// TwinCAT 3 PLC project ExamplePLC
// ProgramVersion: 3.1.4024.0
// libraries:
//   MachineLibrary, * (PLC-Template)
//   Tc2_Standard, * (Beckhoff Automation GmbH)
//   Tc2_System, * (Beckhoff Automation GmbH)
//   Tc2_Utilities, * (Beckhoff Automation GmbH)
//   Tc3_IotBase, * (Beckhoff Automation GmbH)
//   Tc3_JsonXml, * (Beckhoff Automation GmbH)
//   Tc3_Module, * (Beckhoff Automation GmbH)
//   MachineLibrary, * (PLC-Template)
// project tree:
//   Communication/MQTT/_DUTs/ ST_MqttConfiguration.TcDUT, ST_MqttStatus.TcDUT
//   Communication/MQTT/ FB_MqttStatePublisher.TcPOU
//   / PlcTask.TcTTO
//   POUs/ FB_Machine.TcPOU, MAIN.TcPOU
//   Stations/ExampleStation/_DUTs/ ST_ExampleStationConfiguration.TcDUT, ST_ExampleStationStatus.TcDUT
//   Stations/ExampleStation/_ENUMs/ E_ExampleStationRunStep.TcDUT
//   Stations/ExampleStation/ FB_ExampleStation.TcPOU
//   Simulation/SoftwareSim/_DUTs/ ST_ExampleSoftwareSimConfiguration.TcDUT, ST_ExampleSoftwareSimStatus.TcDUT
//   Simulation/SoftwareSim/_ENUMs/ E_ExampleSoftwareSimStep.TcDUT
//   Simulation/SoftwareSim/ FB_ExampleSoftwareSim.TcPOU
//   Stations/ExampleStation/Transaction/_DUTs/ ST_ExampleRequest.TcDUT, ST_ExampleResponse.TcDUT
//   Stations/ExampleStation/Transaction/ FB_ExampleTransaction.TcPOU
//   Simulation/DosingProcessSim/_DUTs/ ST_DosingProcessSimConfiguration.TcDUT, ST_DosingProcessSimStatus.TcDUT
//   Simulation/DosingProcessSim/ FB_DosingProcessSim.TcPOU
//   Stations/DosingStation/_DUTs/ ST_DosingStationConfiguration.TcDUT, ST_DosingStationStatus.TcDUT
//   Stations/DosingStation/ FB_DosingStation.TcPOU
// real-time tasks:
//   TASK PlcTask: cycle T#10ms, priority 20, ADS port 350

CONFIGURATION ExamplePLC
    RESOURCE PLC ON TwinCAT3
        TASK PlcTask(INTERVAL := T#10ms, PRIORITY := 20);
        PROGRAM MAIN WITH PlcTask : MAIN;
    END_RESOURCE
END_CONFIGURATION

// ---- Communication/MQTT/_DUTs/ST_MqttConfiguration.TcDUT
TYPE ST_MqttConfiguration :
STRUCT
	enable					: BOOL := TRUE; //connect to the broker and publish state
	hostName				: STRING(255) := 'broker.hivemq.com'; //public test broker, replace with your own
	hostPort				: UINT := 1883; //8883 for TLS
	stateTopic				: STRING(255) := 'plc-template/example/state'; //machine state is published here as JSON
	commandTopic			: STRING(255) := 'plc-template/example/cmd'; //START, STOP or RESET
	enableRemoteCommands	: BOOL := FALSE; //accept commands on commandTopic. Off by default: anyone on a public broker can publish to it
	publishInterval			: TIME := T#10S; //state is also published on every state change
END_STRUCT
END_TYPE

// ---- Communication/MQTT/_DUTs/ST_MqttStatus.TcDUT
TYPE ST_MqttStatus :
STRUCT
	connected				: BOOL; //connected to the broker
	subscribed				: BOOL; //subscribed to commandTopic
	error					: BOOL; //client error
	errorCode				: HRESULT; //client error code
	publishCount			: UDINT; //messages published
	lastPayloadIn			: STRING(255); //last payload received on commandTopic
END_STRUCT
END_TYPE

// ---- Stations/ExampleStation/_DUTs/ST_ExampleStationConfiguration.TcDUT
TYPE ST_ExampleStationConfiguration :
STRUCT
	cycleDwell			: TIME := T#2S; //wait time between jobs while running
	maxCloseDwell		: TIME := T#10S; //longest closeDwell accepted in a request
END_STRUCT
END_TYPE

// ---- Stations/ExampleStation/_DUTs/ST_ExampleStationStatus.TcDUT
TYPE ST_ExampleStationStatus :
STRUCT
	runStep				: E_ExampleStationRunStep := E_ExampleStationRunStep.Idle; //running sequence step
	allOpen				: BOOL; //both actuators at home (open)
	allClosed			: BOOL; //both actuators at work (closed)
	
	job					: ST_ExampleRequest; //job being worked on
	cycleCount			: UDINT; //completed jobs
	lastCycleTime		: TIME; //duration of the last close/hold/open cycle
	jobsRejected		: UDINT; //requests rejected as invalid
	lastRejectText		: T_MaxString; //reason for the last rejection
	commError			: BOOL; //transaction timed out waiting for the software
END_STRUCT
END_TYPE

// ---- Stations/ExampleStation/_ENUMs/E_ExampleStationRunStep.TcDUT
{attribute 'qualified_only'}
{attribute 'strict'}
{attribute 'to_string'}
TYPE E_ExampleStationRunStep :
(
	Idle			:= 0, //not running
	RequestJob		:= 10, //raise attention, ask the software for a job
	WaitJob			:= 20, //wait for the request, validate it, ack or reject
	WaitWorking		:= 30, //wait for the software to drop trigger
	Close			:= 40, //closing both actuators
	HoldClosed		:= 50, //holding closed for the requested closeDwell
	Open			:= 60, //opening both actuators
	Report			:= 70, //send the response with tell
	WaitReportAck	:= 80, //wait for the software to acknowledge the response
	Dwell			:= 90 //wait before requesting the next job
);
END_TYPE

// ---- Simulation/SoftwareSim/_DUTs/ST_ExampleSoftwareSimConfiguration.TcDUT
TYPE ST_ExampleSoftwareSimConfiguration :
STRUCT
	enable				: BOOL := TRUE; //answer the station's transactions
	responseDelay		: TIME := T#500MS; //delay before each software action
	closeDwell			: TIME := T#1S; //closeDwell sent in each request
	
	//Fault injection
	freeze				: BOOL; //stop responding where it is (tests the commTimeout)
	sendInvalidRequest	: BOOL; //send closeDwell = T#0S (station should reject it)
END_STRUCT
END_TYPE

// ---- Simulation/SoftwareSim/_DUTs/ST_ExampleSoftwareSimStatus.TcDUT
TYPE ST_ExampleSoftwareSimStatus :
STRUCT
	step				: E_ExampleSoftwareSimStep := E_ExampleSoftwareSimStep.Idle; //current step
	requestsSent		: UDINT; //requests sent (trigger raised)
	responsesReceived	: UDINT; //responses received (tell acknowledged)
	aborts				: UDINT; //transactions aborted by the PLC
	lastResponse		: ST_ExampleResponse; //last response read on tell
END_STRUCT
END_TYPE

// ---- Simulation/SoftwareSim/_ENUMs/E_ExampleSoftwareSimStep.TcDUT
{attribute 'qualified_only'}
{attribute 'strict'}
{attribute 'to_string'}
TYPE E_ExampleSoftwareSimStep :
(
	Idle			:= 0, //waiting for attention
	SendTrigger		:= 10, //delay, then raise trigger with a request
	WaitTriggerAck	:= 20, //waiting for trigger_ack
	DropTrigger		:= 30, //delay, then drop trigger
	WaitTell		:= 40, //waiting for tell
	SendTellAck		:= 50, //delay, read response, raise tell_ack
	WaitTellDrop	:= 60, //waiting for tell to drop
	DropTellAck		:= 70 //drop tell_ack, transaction closed
);
END_TYPE

// ---- Stations/ExampleStation/Transaction/_DUTs/ST_ExampleRequest.TcDUT
(* Request from the software to the station, sent with trigger. *)
TYPE ST_ExampleRequest :
STRUCT
	cycleId				: UDINT; //id chosen by the software, echoed back in the response
	closeDwell			: TIME; //how long to hold the actuators closed
END_STRUCT
END_TYPE

// ---- Stations/ExampleStation/Transaction/_DUTs/ST_ExampleResponse.TcDUT
(* Response from the station to the software, sent with tell. *)
TYPE ST_ExampleResponse :
STRUCT
	cycleId				: UDINT; //cycleId from the request
	cycleTime			: TIME; //time to close, hold and open
	ok					: BOOL; //cycle completed without faults
END_STRUCT
END_TYPE

// ---- Simulation/DosingProcessSim/_DUTs/ST_DosingProcessSimConfiguration.TcDUT
TYPE ST_DosingProcessSimConfiguration :
STRUCT
	enable				: BOOL := TRUE; //simulate the flows (turn off when real I/O is linked)
	mainFlowBase		: LREAL := 200; //average main flow in l/min (set below 50 to test the low-low interlock)
	mainFlowSwing		: LREAL := 50; //main flow varies +/- this much in l/min
	swingPeriod			: TIME := T#60S; //period of the main flow variation, T#0S = constant
	maxDosingFlow		: LREAL := 80; //dosing flow at 100 % valve in l/min
	processLag			: TIME := T#2S; //time constant from valve position to dosing flow
END_STRUCT
END_TYPE

// ---- Simulation/DosingProcessSim/_DUTs/ST_DosingProcessSimStatus.TcDUT
TYPE ST_DosingProcessSimStatus :
STRUCT
	mainFlow			: LREAL; //simulated main flow in l/min
	dosingFlow			: LREAL; //simulated dosing flow in l/min
END_STRUCT
END_TYPE

// ---- Stations/DosingStation/_DUTs/ST_DosingStationConfiguration.TcDUT
TYPE ST_DosingStationConfiguration :
STRUCT
	ratio				: LREAL := 0.2; //dosing flow / main flow while running
END_STRUCT
END_TYPE

// ---- Stations/DosingStation/_DUTs/ST_DosingStationStatus.TcDUT
TYPE ST_DosingStationStatus :
STRUCT
	dosing				: BOOL; //PID in ratio control
	mainFlow			: LREAL; //main flow in l/min
	dosingFlow			: LREAL; //dosing flow in l/min
	dosingSetpoint		: LREAL; //dosing flow setpoint from the ratio, in l/min
	ratioActual			: LREAL; //dosing flow / main flow
	valvePosition		: LREAL; //dosing valve position in %
	mainFlowLow			: BOOL; //main flow below its low-low limit: dosing valve interlocked closed
END_STRUCT
END_TYPE

// ---- POUs/MAIN.TcPOU
PROGRAM MAIN
VAR
	{attribute 'OPC.UA.DA' := '1'}
	machine		: FB_Machine; //top-level module, start/stop with machine.ocmd
	
	(* Test harness
	----------------------------------------------------------------------------------------------------*)
	{attribute 'OPC.UA.DA' := '1'}
	softwareSim	: FB_ExampleSoftwareSim; //plays the software side of the station's trigger/tell
	{attribute 'OPC.UA.DA' := '1'}
	dosingSim	: FB_DosingProcessSim; //simulates the dosing station's flows
END_VAR

machine();

//Outside world: answers the example station's job requests
softwareSim(transaction := machine.exampleStation.transaction);

//Process simulation for the dosing station (turn off with dosingSim.cfg.enable when I/O is linked)
dosingSim(station := machine.dosingStation);

END_PROGRAM

// ---- POUs/FB_Machine.TcPOU
FUNCTION_BLOCK FB_Machine EXTENDS FB_Module
(*
	Top-level module. Starting/stopping the machine starts/stops both stations.
	Start/stop/reset from the HMI with ocmd, or over MQTT (see cfgMqtt.enableRemoteCommands).
*)
VAR_INPUT
	(* Stations
	----------------------------------------------------------------------------------------------------*)
	{attribute 'OPC.UA.DA' := '1'}
	exampleStation		: FB_ExampleStation;
	{attribute 'OPC.UA.DA' := '1'}
	dosingStation		: FB_DosingStation; //ratio control loop example
	
	(* Communication
	----------------------------------------------------------------------------------------------------*)
	{attribute 'OPC.UA.DA' := '1'}
	{attribute 'OPC.UA.DA.StructuredType' := '1'}
	cfgMqtt				: ST_MqttConfiguration; //MQTT configuration
END_VAR
VAR
	{attribute 'OPC.UA.DA' := '0'} // internal MQTT client holds pointers OPC UA can't publish; status is in cfgMqtt/dashboard
	mqtt				: FB_MqttStatePublisher; //MQTT state publisher
END_VAR

SUPER^();

Stations();
Permissives();
Communication();

METHOD PROTECTED Communication
mqtt(cfg 			:= cfgMqtt,
	 machineState 	:= sts.State,
	 cycleCount 	:= exampleStation.stsStation.cycleCount);

//Remote commands are handled like program commands
IF mqtt.cmd <> E_ModuleCommand.None THEN
	pcmd := mqtt.cmd;
END_IF
END_METHOD

METHOD PROTECTED Permissives //set module permissives and interlocks
//Started once every station is running
PermStartComplete.cfg.condText[0] := 'Example station started';
PermStartComplete.cfg.condText[1] := 'Dosing station started';
PermStartComplete.perm.0 := exampleStation.sts.Started;
PermStartComplete.perm.1 := dosingStation.sts.Started;

//Stopped once every station is stopped
PermStopComplete.cfg.condText[0] := 'Example station stopped';
PermStopComplete.cfg.condText[1] := 'Dosing station stopped';
PermStopComplete.perm.0 := exampleStation.sts.Stopped;
PermStopComplete.perm.1 := dosingStation.sts.Stopped;

//A faulted station stops the machine
IntlkAuto.cfg.condText[0] := 'Example station not faulted';
IntlkAuto.cfg.condText[1] := 'Dosing station not faulted';
IntlkAuto.perm.0 := NOT exampleStation.sts.Faulted;
IntlkAuto.perm.1 := NOT dosingStation.sts.Faulted;
END_METHOD

METHOD PUBLIC Reset : BOOL
exampleStation.cmdReset := TRUE;
dosingStation.cmdReset := TRUE;
Reset := TRUE;
END_METHOD

METHOD PROTECTED Started : BOOL
//Stations run their own sequences while the machine is started
END_METHOD

METHOD PROTECTED Starting : BOOL
exampleStation.pcmd := E_ModuleCommand.Start;
dosingStation.pcmd := E_ModuleCommand.Start;
END_METHOD

METHOD PROTECTED Stations //call child modules
exampleStation();
dosingStation();

inpChildFaulted := exampleStation.sts.Faulted OR dosingStation.sts.Faulted;
END_METHOD

METHOD PROTECTED Stopping : BOOL
exampleStation.pcmd := E_ModuleCommand.Stop;
dosingStation.pcmd := E_ModuleCommand.Stop;
END_METHOD

END_FUNCTION_BLOCK

// ---- Stations/ExampleStation/FB_ExampleStation.TcPOU
FUNCTION_BLOCK FB_ExampleStation EXTENDS FB_Module
(*
	Example station with two 2-state actuators and a trigger/tell transaction.
	Home position = OPEN, Work position = CLOSED.
	
	Starting (homing)	: open both actuators, Started once both are open
	Started (running)	: one job per cycle:
						  ask the software for a job (attention), validate and ack the request,
						  close both, hold for request.closeDwell, open both, report (tell), dwell
	Stopping			: abort any open transaction, open both actuators (safe position)
	Stopped				: actuators follow operator commands (manual mode)
	
	The actuators are configured with no feedback so the example runs without hardware.
	Clear homeNoFdbk/workNoFdbk and link homeFdbk/workFdbk/outHome/outWork to use real I/O.
*)
VAR_INPUT
	{attribute 'OPC.UA.DA' := '1'}
	{attribute 'OPC.UA.DA.StructuredType' := '1'}
	cfg					: ST_ExampleStationConfiguration; //configuration
	
	(* Devices
	----------------------------------------------------------------------------------------------------*)
	{attribute 'OPC.UA.DA' := '1'}
	actuatorA			: FB_Actuator2State := (cfg := (actuatorId := 'Actuator A', homeNoFdbk := TRUE, workNoFdbk := TRUE));
	{attribute 'OPC.UA.DA' := '1'}
	actuatorB			: FB_Actuator2State := (cfg := (actuatorId := 'Actuator B', homeNoFdbk := TRUE, workNoFdbk := TRUE));
	
	(* Communication
	----------------------------------------------------------------------------------------------------*)
	{attribute 'OPC.UA.DA' := '1'}
	transaction			: FB_ExampleTransaction := (cfg := (commTimeout := T#10S)); //job request/response with the software
END_VAR
VAR_OUTPUT
	{attribute 'OPC.UA.DA' := '1'}
	{attribute 'OPC.UA.DA.Access' := '1'}
	{attribute 'OPC.UA.DA.StructuredType' := '1'}
	stsStation			: ST_ExampleStationStatus; //station specific status (module status is in sts)
END_VAR
VAR
	//Timers
	dwellTimer			: TON; //dwell between cycles
	holdTimer			: TON; //holds the actuators closed for job.closeDwell
	cycleTimer			: TON := (PT := T#1D); //measures one close/hold/open cycle
END_VAR

SUPER^();

Devices();
Permissives();
StatusOut();

METHOD PROTECTED CloseAll //command all actuators to work (closed)
IF NOT actuatorA.sts.atWork AND NOT actuatorA.sts.goingToWork THEN
	actuatorA.ToWork();
END_IF
IF NOT actuatorB.sts.atWork AND NOT actuatorB.sts.goingToWork THEN
	actuatorB.ToWork();
END_IF
END_METHOD

METHOD PROTECTED Devices //call child devices
//Devices follow this module's mode through childCtrl
actuatorA(parentCtrl := childCtrl);
actuatorB(parentCtrl := childCtrl);
transaction();

//Report child faults to the module
inpChildFaulted := actuatorA.fault.active OR actuatorB.fault.active;
END_METHOD

METHOD PROTECTED OpenAll //command all actuators to home (open)
IF NOT actuatorA.sts.atHome AND NOT actuatorA.sts.goingToHome THEN
	actuatorA.ToHome();
END_IF
IF NOT actuatorB.sts.atHome AND NOT actuatorB.sts.goingToHome THEN
	actuatorB.ToHome();
END_IF
END_METHOD

METHOD PROTECTED Permissives //set module permissives and interlocks
//Homing is complete when all actuators are open
PermStartComplete.cfg.condText[0] := 'Actuator A open';
PermStartComplete.cfg.condText[1] := 'Actuator B open';
PermStartComplete.perm.0 := actuatorA.sts.atHome;
PermStartComplete.perm.1 := actuatorB.sts.atHome;

//Stopping is complete when all actuators are open, or faulted so they cannot move
PermStopComplete.cfg.condText[0] := 'Actuator A open or faulted';
PermStopComplete.cfg.condText[1] := 'Actuator B open or faulted';
PermStopComplete.perm.0 := actuatorA.sts.atHome OR actuatorA.fault.active;
PermStopComplete.perm.1 := actuatorB.sts.atHome OR actuatorB.fault.active;

//A faulted actuator stops the station
IntlkAuto.cfg.condText[0] := 'Actuator A not faulted';
IntlkAuto.cfg.condText[1] := 'Actuator B not faulted';
IntlkAuto.perm.0 := NOT actuatorA.fault.active;
IntlkAuto.perm.1 := NOT actuatorB.fault.active;
END_METHOD

METHOD PUBLIC Reset : BOOL
actuatorA.Reset();
actuatorB.Reset();
transaction.Reset();
Reset := TRUE;
END_METHOD

METHOD PROTECTED Started : BOOL
//Running sequence: one trigger/tell transaction per close/open cycle
CASE stsStation.runStep OF
	
	E_ExampleStationRunStep.Idle:
		stsStation.runStep := E_ExampleStationRunStep.RequestJob;
		
	E_ExampleStationRunStep.RequestJob:
		IF transaction.sts.Idle THEN
			transaction.Start(); //raises attention
			stsStation.runStep := E_ExampleStationRunStep.WaitJob;
		END_IF
		
	E_ExampleStationRunStep.WaitJob:
		IF transaction.sts.Request_Start THEN
			IF ValidateJob(transaction.request) THEN
				stsStation.job := transaction.request;
				transaction.SetRequestACK();
				stsStation.runStep := E_ExampleStationRunStep.WaitWorking;
			ELSE
				transaction.Abort();
				stsStation.jobsRejected := stsStation.jobsRejected + 1;
				stsStation.runStep := E_ExampleStationRunStep.Dwell;
			END_IF
		END_IF
		
	E_ExampleStationRunStep.WaitWorking:
		IF transaction.sts.Working THEN
			stsStation.runStep := E_ExampleStationRunStep.Close;
		END_IF
		
	E_ExampleStationRunStep.Close:
		CloseAll();
		IF stsStation.allClosed THEN
			stsStation.runStep := E_ExampleStationRunStep.HoldClosed;
		END_IF
		
	E_ExampleStationRunStep.HoldClosed:
		IF holdTimer.Q THEN
			stsStation.runStep := E_ExampleStationRunStep.Open;
		END_IF
		
	E_ExampleStationRunStep.Open:
		OpenAll();
		IF stsStation.allOpen THEN
			stsStation.lastCycleTime := cycleTimer.ET;
			stsStation.runStep := E_ExampleStationRunStep.Report;
		END_IF
		
	E_ExampleStationRunStep.Report:
		transaction.response.cycleId 	:= stsStation.job.cycleId;
		transaction.response.cycleTime 	:= stsStation.lastCycleTime;
		transaction.response.ok 		:= NOT (actuatorA.fault.active OR actuatorB.fault.active);
		transaction.FinishWork(); //raises tell
		stsStation.cycleCount := stsStation.cycleCount + 1;
		stsStation.runStep := E_ExampleStationRunStep.WaitReportAck;
		
	E_ExampleStationRunStep.WaitReportAck:
		IF transaction.sts.Idle THEN
			stsStation.runStep := E_ExampleStationRunStep.Dwell;
		END_IF
		
	E_ExampleStationRunStep.Dwell:
		IF dwellTimer.Q THEN
			stsStation.runStep := E_ExampleStationRunStep.RequestJob;
		END_IF
		
END_CASE
END_METHOD

METHOD PROTECTED Starting : BOOL
//Homing: open all actuators, no transaction open
OpenAll();
AbortTransaction();
stsStation.runStep := E_ExampleStationRunStep.Idle;
END_METHOD

METHOD PROTECTED StatusOut //Set output status information
stsStation.allOpen 	:= actuatorA.sts.atHome AND actuatorB.sts.atHome;
stsStation.allClosed 	:= actuatorA.sts.atWork AND actuatorB.sts.atWork;

stsStation.commError 	:= transaction.sts.errTimeout;

//Monitoring timers
dwellTimer(IN := stsStation.runStep = E_ExampleStationRunStep.Dwell, PT := cfg.cycleDwell);
holdTimer(IN := stsStation.runStep = E_ExampleStationRunStep.HoldClosed, PT := stsStation.job.closeDwell);
cycleTimer(IN := stsStation.runStep = E_ExampleStationRunStep.Close
			OR stsStation.runStep = E_ExampleStationRunStep.HoldClosed
			OR stsStation.runStep = E_ExampleStationRunStep.Open);
END_METHOD

METHOD PROTECTED Stopping : BOOL
//Finish in the safe position: all actuators open, transaction closed
OpenAll();
AbortTransaction();
stsStation.runStep := E_ExampleStationRunStep.Idle;
END_METHOD

METHOD PROTECTED AbortTransaction //cancel an open transaction
IF transaction.sts.bBusy THEN
	transaction.Abort();
END_IF
END_METHOD

METHOD PROTECTED ValidateJob : BOOL //TRUE if the request can be worked on, sets lastRejectText otherwise
VAR_INPUT
	job			: ST_ExampleRequest;
END_VAR
IF job.closeDwell <= T#0S THEN
	stsStation.lastRejectText := 'closeDwell must be greater than 0';
ELSIF job.closeDwell > cfg.maxCloseDwell THEN
	stsStation.lastRejectText := 'closeDwell is longer than cfg.maxCloseDwell';
ELSE
	ValidateJob := TRUE;
	RETURN;
END_IF
ValidateJob := FALSE;
END_METHOD

END_FUNCTION_BLOCK

// ---- Stations/ExampleStation/Transaction/FB_ExampleTransaction.TcPOU
FUNCTION_BLOCK FB_ExampleTransaction EXTENDS FB_TriggerTell
(*
	Trigger/tell transaction for the example station, carrying ST_ExampleRequest in
	and ST_ExampleResponse out.
	
	FB_TriggerTell keeps its handshake bits internal. This FB is the transport layer:
	the software side writes trigger/tell_ack with WriteTrigger()/WriteTellAck() and
	reads the PLC bits from handshake. A real project would map these to OPC UA or MQTT.
*)
VAR_INPUT
	{attribute 'OPC.UA.DA' := '1'}
	{attribute 'OPC.UA.DA.StructuredType' := '1'}
	response			: ST_ExampleResponse; //set by the station before FinishWork()
END_VAR
VAR_OUTPUT
	{attribute 'OPC.UA.DA' := '1'}
	{attribute 'OPC.UA.DA.Access' := '1'}
	{attribute 'OPC.UA.DA.StructuredType' := '1'}
	request				: ST_ExampleRequest; //request latched when trigger rises
	{attribute 'OPC.UA.DA' := '1'}
	{attribute 'OPC.UA.DA.Access' := '1'}
	{attribute 'OPC.UA.DA.StructuredType' := '1'}
	handshake			: ST_TriggerTellHandshake; //copy of all handshake bits for the software side
END_VAR
VAR
	requestIn			: ST_ExampleRequest; //request written by the software with trigger
	
	//Oneshot triggers
	rtTrigger			: R_TRIG;
END_VAR

//Latch the request when the software raises trigger
rtTrigger(CLK := stHandshake.trigger);
IF rtTrigger.Q THEN
	request := requestIn;
END_IF

SUPER^();

handshake := stHandshake;

METHOD PUBLIC Response_Cleanup : BOOL //clear the response once the software acknowledged it
VAR
	emptyResponse : ST_ExampleResponse;
END_VAR
SUPER^.Response_Cleanup();
response := emptyResponse;
Response_Cleanup := TRUE;
END_METHOD

METHOD PUBLIC WriteTellAck //software side: set or clear tell_ack
VAR_INPUT
	value		: BOOL;
END_VAR
stHandshake.tell_ack := value;
END_METHOD

METHOD PUBLIC WriteTrigger //software side: set or clear trigger, with the request data
VAR_INPUT
	value		: BOOL;
	req			: ST_ExampleRequest; //only used when value is TRUE
END_VAR
IF value THEN
	requestIn := req;
END_IF
stHandshake.trigger := value;
END_METHOD

END_FUNCTION_BLOCK

// ---- Stations/DosingStation/FB_DosingStation.TcPOU
FUNCTION_BLOCK FB_DosingStation EXTENDS FB_Module
(*
	Example of a ratio control loop built from MachineLibrary blocks:
	
		flowMain (FB_AnalogInput)	main flow, the "wild" flow nobody controls
		flowDosing (FB_AnalogInput)	dosing flow, the process value
		dosingPid (FB_PID)			Ratio mode: dosing setpoint = cfg.ratio x main flow
		dosingValve					FB_ActuatorModulating driven by the PID output
	
	Starting	: PID off, valve closed
	Started		: PID in Ratio mode at cfg.ratio
	Stopping	: PID off, valve closed
	Interlock	: main flow low-low closes the valve (dosing into no flow is unsafe)
	
	No hardware needed: the valve has no position feedback (simulated stroke) and
	MAIN.dosingSim writes both flows into the analog inputs' simulation values.
	For real I/O, link flowMain.inpRaw, flowDosing.inpRaw and dosingValve.outRaw,
	and turn off MAIN.dosingSim.
*)
VAR_INPUT
	{attribute 'OPC.UA.DA' := '1'}
	{attribute 'OPC.UA.DA.StructuredType' := '1'}
	cfg					: ST_DosingStationConfiguration; //configuration
	
	(* Devices
	----------------------------------------------------------------------------------------------------*)
	{attribute 'OPC.UA.DA' := '1'}
	flowMain			: FB_AnalogInput := (cfg := (inputId := 'Main flow', units := 'l/min', euMax := 400, filterTime := T#500MS, limits := (LowLow := 50, Low := 100, High := 350, HighHigh := 380), alarmEnable := (lowLow := TRUE, low := TRUE, high := TRUE, highHigh := TRUE)));
	{attribute 'OPC.UA.DA' := '1'}
	flowDosing			: FB_AnalogInput := (cfg := (inputId := 'Dosing flow', units := 'l/min', euMax := 100, filterTime := T#500MS));
	{attribute 'OPC.UA.DA' := '1'}
	dosingPid			: FB_PID := (cfg := (loopId := 'Dosing', kp := 1.5, ti := T#3S, setpointMax := 100, ratioMax := 1, deviationEnable := TRUE, deviationLimit := 10));
	{attribute 'OPC.UA.DA' := '1'}
	dosingValve			: FB_ActuatorModulating := (cfg := (actuatorId := 'Dosing valve', noFdbk := TRUE, strokeTime := T#10S, failTimePositioning := T#30S));
END_VAR
VAR_OUTPUT
	{attribute 'OPC.UA.DA' := '1'}
	{attribute 'OPC.UA.DA.Access' := '1'}
	{attribute 'OPC.UA.DA.StructuredType' := '1'}
	stsStation			: ST_DosingStationStatus; //station specific status (module status is in sts)
END_VAR
VAR
END_VAR

SUPER^();

Devices();
Permissives();
StatusOut();

METHOD PROTECTED Devices //call child devices and connect the loop
//Inputs first, so the PID sees this scan's values
flowMain();
flowDosing();

dosingPid(pv		:= flowDosing.sts.value,
		  wildValue	:= flowMain.sts.value,
		  inpPvBad	:= NOT flowDosing.sts.valid,
		  parentCtrl := childCtrl);

//Dosing into a low main flow is not allowed: losing this closes the valve
dosingValve.intlk.cfg.condText[0] := 'Main flow not low-low';
dosingValve.intlk.perm.0 := NOT flowMain.sts.lowLow;
dosingValve(parentCtrl := childCtrl);

//PID output to the valve (program commands are only accepted in Auto)
IF dosingPid.sts.closedLoop AND dosingValve.sts.modeAuto THEN
	dosingValve.SetPosition(dosingPid.out);
END_IF

//Report child faults to the module
inpChildFaulted := dosingValve.fault.active OR dosingPid.fault.active
				OR flowMain.fault.active OR flowDosing.fault.active;
END_METHOD

METHOD PROTECTED Permissives //set module permissives and interlocks
//Homing is complete when the valve is closed and the loop is off
PermStartComplete.cfg.condText[0] := 'Dosing valve closed';
PermStartComplete.cfg.condText[1] := 'Dosing loop off';
PermStartComplete.perm.0 := dosingValve.sts.closed;
PermStartComplete.perm.1 := dosingPid.sts.loopMode = E_PIDLoopMode.Off;

//Stopping is complete when the valve is closed, or faulted so it cannot move
PermStopComplete.cfg.condText[0] := 'Dosing valve closed or faulted';
PermStopComplete.perm.0 := dosingValve.sts.closed OR dosingValve.fault.active;

//Faults stop the station
IntlkAuto.cfg.condText[0] := 'Dosing valve not faulted';
IntlkAuto.cfg.condText[1] := 'Dosing loop not faulted';
IntlkAuto.cfg.condText[2] := 'Flow signals good';
IntlkAuto.perm.0 := NOT dosingValve.fault.active;
IntlkAuto.perm.1 := NOT dosingPid.fault.active;
IntlkAuto.perm.2 := NOT (flowMain.fault.active OR flowDosing.fault.active);
END_METHOD

METHOD PUBLIC Reset : BOOL
flowMain.Reset();
flowDosing.Reset();
dosingPid.Reset();
dosingValve.Reset();
Reset := TRUE;
END_METHOD

METHOD PROTECTED Started : BOOL
//Running: ratio control. Re-issued when the ratio changes.
IF dosingPid.sts.loopMode <> E_PIDLoopMode.Ratio OR dosingPid.sts.ratio <> cfg.ratio THEN
	dosingPid.Ratio(cfg.ratio);
END_IF
END_METHOD

METHOD PROTECTED Starting : BOOL
//Homing: loop off, valve closed
SafeState();
END_METHOD

METHOD PROTECTED Stopping : BOOL
//Finish in the safe state: loop off, valve closed
SafeState();
END_METHOD

METHOD PROTECTED SafeState //loop off and valve closed
IF dosingPid.sts.loopMode <> E_PIDLoopMode.Off THEN
	dosingPid.Off();
END_IF
IF NOT dosingValve.sts.closed AND dosingValve.sts.setpoint <> dosingValve.cfg.minPosition THEN
	dosingValve.Close();
END_IF
END_METHOD

METHOD PROTECTED StatusOut //Set output status information
stsStation.dosing			:= dosingPid.sts.loopMode = E_PIDLoopMode.Ratio;
stsStation.mainFlow			:= flowMain.sts.value;
stsStation.dosingFlow		:= flowDosing.sts.value;
stsStation.dosingSetpoint	:= dosingPid.sts.setpoint;
stsStation.valvePosition	:= dosingValve.sts.position;
stsStation.mainFlowLow		:= flowMain.sts.lowLow;
IF flowMain.sts.value > 0 THEN
	stsStation.ratioActual := flowDosing.sts.value / flowMain.sts.value;
ELSE
	stsStation.ratioActual := 0;
END_IF
END_METHOD

END_FUNCTION_BLOCK

// ---- Communication/MQTT/FB_MqttStatePublisher.TcPOU
FUNCTION_BLOCK FB_MqttStatePublisher
(*
	Publishes the machine state as JSON over MQTT, and optionally accepts START/STOP/RESET.
	Shows how Tc3_IotBase and Tc3_JsonXml are used next to MachineLibrary.
	Payload example: {"state":"Started","cycleCount":12}
*)
VAR_INPUT
	{attribute 'OPC.UA.DA' := '1'}
	{attribute 'OPC.UA.DA.StructuredType' := '1'}
	cfg					: ST_MqttConfiguration; //configuration
	
	machineState		: E_ModuleState; //state to publish
	cycleCount			: UDINT; //cycle count to publish
END_VAR
VAR_OUTPUT
	cmd					: E_ModuleCommand; //remote command received this scan, None otherwise
	
	{attribute 'OPC.UA.DA' := '1'}
	{attribute 'OPC.UA.DA.Access' := '1'}
	{attribute 'OPC.UA.DA.StructuredType' := '1'}
	sts					: ST_MqttStatus;
END_VAR
VAR
	bInit				: BOOL := TRUE;
	
	//MQTT client
	client				: FB_IotMqttClient;
	queue				: FB_IotMqttMessageQueue;
	message				: FB_IotMqttMessage;
	
	//Publish
	json				: FB_JsonSaxWriter;
	stateText			: STRING;
	payloadOut			: STRING(255);
	publishRequest		: BOOL;
	machineStateLast	: E_ModuleState := E_ModuleState.Unknown;
	publishTimer		: TON;
	
	//Subscribe
	{attribute 'TcEncoding' := 'UTF-8'}
	topicIn				: STRING(255);
	{attribute 'TcEncoding' := 'UTF-8'}
	payloadIn			: STRING(255);
END_VAR

cmd := E_ModuleCommand.None;

IF NOT cfg.enable THEN
	sts.connected := sts.subscribed := FALSE;
	RETURN;
END_IF

IF bInit THEN
	Init();
	bInit := FALSE;
END_IF

Connection();
Publish();
Subscribe();

METHOD PROTECTED Connection //keep the client connected (must run every scan)
client.Execute(bConnect := TRUE);

sts.connected 	:= client.bConnected;
sts.error 		:= client.bError;
sts.errorCode 	:= client.hrErrorCode;
END_METHOD

METHOD PROTECTED Init : BOOL
client.sHostName 		:= cfg.hostName;
client.nHostPort 		:= cfg.hostPort;
client.ipMessageQueue 	:= queue; //route received messages into the queue
Init := TRUE;
END_METHOD

METHOD PROTECTED Publish //publish on state change and every publishInterval
publishTimer(IN := sts.connected AND NOT publishTimer.Q, PT := cfg.publishInterval);
publishRequest := publishRequest OR publishTimer.Q OR (machineState <> machineStateLast);
machineStateLast := machineState;

IF publishRequest AND sts.connected THEN
	stateText := TO_STRING(machineState);
	
	json.ResetDocument();
	json.StartObject();
	json.AddKey('state');
	json.AddString(stateText);
	json.AddKey('cycleCount');
	json.AddDint(UDINT_TO_DINT(cycleCount));
	json.EndObject();
	json.CopyDocument(payloadOut, SIZEOF(payloadOut));
	
	IF client.Publish(
		sTopic			:= cfg.stateTopic,
		pPayload		:= ADR(payloadOut),
		nPayloadSize	:= INT_TO_UDINT(LEN(payloadOut)),
		eQoS			:= TcIotMqttQos.AtMostOnceDelivery,
		bRetain			:= FALSE,
		bQueue			:= FALSE)
	THEN
		publishRequest := FALSE;
		sts.publishCount := sts.publishCount + 1;
	END_IF
END_IF
END_METHOD

METHOD PROTECTED Subscribe //receive remote commands
IF NOT cfg.enableRemoteCommands THEN
	RETURN;
END_IF

IF sts.connected AND NOT sts.subscribed THEN
	sts.subscribed := client.Subscribe(sTopic := cfg.commandTopic, eQoS := TcIotMqttQos.AtMostOnceDelivery);
ELSIF NOT sts.connected THEN
	sts.subscribed := FALSE;
END_IF

IF queue.nQueuedMessages > 0 THEN
	IF queue.Dequeue(fbMessage := message) THEN
		MEMSET(ADR(payloadIn), 0, SIZEOF(payloadIn));
		message.GetTopic(pTopic := ADR(topicIn), nTopicSize := SIZEOF(topicIn));
		message.GetPayload(pPayload := ADR(payloadIn), nPayloadSize := SIZEOF(payloadIn), bSetNullTermination := TRUE);
		sts.lastPayloadIn := payloadIn;
		
		IF payloadIn = 'START' THEN
			cmd := E_ModuleCommand.Start;
		ELSIF payloadIn = 'STOP' THEN
			cmd := E_ModuleCommand.Stop;
		ELSIF payloadIn = 'RESET' THEN
			cmd := E_ModuleCommand.Reset;
		END_IF
	END_IF
END_IF
END_METHOD

END_FUNCTION_BLOCK

// ---- Simulation/SoftwareSim/FB_ExampleSoftwareSim.TcPOU
FUNCTION_BLOCK FB_ExampleSoftwareSim
(*
	Plays the software (MES) side of FB_ExampleTransaction so the trigger/tell
	handshake can be tested without any outside software.
	
	For each transaction: wait for attention, send a request with trigger, drop trigger
	after trigger_ack, read the response on tell, acknowledge with tell_ack.
	Use cfg.freeze and cfg.sendInvalidRequest to test timeouts and rejected requests.
*)
VAR_INPUT
	{attribute 'OPC.UA.DA' := '1'}
	{attribute 'OPC.UA.DA.StructuredType' := '1'}
	cfg					: ST_ExampleSoftwareSimConfiguration; //configuration
END_VAR
VAR_IN_OUT
	transaction			: FB_ExampleTransaction; //transaction to answer
END_VAR
VAR_OUTPUT
	{attribute 'OPC.UA.DA' := '1'}
	{attribute 'OPC.UA.DA.Access' := '1'}
	{attribute 'OPC.UA.DA.StructuredType' := '1'}
	sts					: ST_ExampleSoftwareSimStatus;
END_VAR
VAR
	request				: ST_ExampleRequest; //request being sent
	nextCycleId			: UDINT; //last cycleId sent
	
	//state variables for tracking
	stepLastScan		: E_ExampleSoftwareSimStep;
	
	//Timers
	delayTimer			: TON; //responseDelay, restarts on every step change
END_VAR

IF NOT cfg.enable THEN
	RETURN;
END_IF

HandleAbort();
StateMachine();

METHOD PROTECTED HandleAbort //PLC aborted mid-transaction: drop our bits and start over
IF transaction.sts.Idle AND sts.step >= E_ExampleSoftwareSimStep.WaitTriggerAck THEN
	transaction.WriteTrigger(value := FALSE, req := request);
	transaction.WriteTellAck(value := FALSE);
	sts.aborts := sts.aborts + 1;
	sts.step := E_ExampleSoftwareSimStep.Idle;
END_IF
END_METHOD

METHOD PROTECTED StateMachine
//Restart the delay on every step change, hold it while frozen
delayTimer(IN := (sts.step = stepLastScan) AND NOT cfg.freeze, PT := cfg.responseDelay);
stepLastScan := sts.step;

IF cfg.freeze THEN
	RETURN;
END_IF

CASE sts.step OF
	
	E_ExampleSoftwareSimStep.Idle:
		IF transaction.handshake.attention THEN
			sts.step := E_ExampleSoftwareSimStep.SendTrigger;
		END_IF
		
	E_ExampleSoftwareSimStep.SendTrigger:
		IF delayTimer.Q THEN
			nextCycleId 		:= nextCycleId + 1;
			request.cycleId 	:= nextCycleId;
			request.closeDwell 	:= SEL(cfg.sendInvalidRequest, cfg.closeDwell, T#0S);
			transaction.WriteTrigger(value := TRUE, req := request);
			sts.requestsSent 	:= sts.requestsSent + 1;
			sts.step 			:= E_ExampleSoftwareSimStep.WaitTriggerAck;
		END_IF
		
	E_ExampleSoftwareSimStep.WaitTriggerAck:
		IF transaction.handshake.trigger_ack THEN
			sts.step := E_ExampleSoftwareSimStep.DropTrigger;
		END_IF
		
	E_ExampleSoftwareSimStep.DropTrigger:
		IF delayTimer.Q THEN
			transaction.WriteTrigger(value := FALSE, req := request);
			sts.step := E_ExampleSoftwareSimStep.WaitTell;
		END_IF
		
	E_ExampleSoftwareSimStep.WaitTell:
		IF transaction.handshake.tell THEN
			sts.step := E_ExampleSoftwareSimStep.SendTellAck;
		END_IF
		
	E_ExampleSoftwareSimStep.SendTellAck:
		IF delayTimer.Q THEN
			sts.lastResponse 		:= transaction.response;
			sts.responsesReceived 	:= sts.responsesReceived + 1;
			transaction.WriteTellAck(value := TRUE);
			sts.step 				:= E_ExampleSoftwareSimStep.WaitTellDrop;
		END_IF
		
	E_ExampleSoftwareSimStep.WaitTellDrop:
		IF NOT transaction.handshake.tell THEN
			sts.step := E_ExampleSoftwareSimStep.DropTellAck;
		END_IF
		
	E_ExampleSoftwareSimStep.DropTellAck:
		transaction.WriteTellAck(value := FALSE);
		sts.step := E_ExampleSoftwareSimStep.Idle;
		
END_CASE
END_METHOD

END_FUNCTION_BLOCK

// ---- Simulation/DosingProcessSim/FB_DosingProcessSim.TcPOU
FUNCTION_BLOCK FB_DosingProcessSim
(*
	Simulates the process behind FB_DosingStation so the loop runs without hardware.
	Main flow swings around cfg.mainFlowBase; dosing flow follows the valve position
	through a first-order lag. Both are written to the analog inputs' simulation values.
*)
VAR_INPUT
	{attribute 'OPC.UA.DA' := '1'}
	{attribute 'OPC.UA.DA.StructuredType' := '1'}
	cfg					: ST_DosingProcessSimConfiguration; //configuration
END_VAR
VAR_IN_OUT
	station				: FB_DosingStation; //station to simulate
END_VAR
VAR_OUTPUT
	{attribute 'OPC.UA.DA' := '1'}
	{attribute 'OPC.UA.DA.Access' := '1'}
	{attribute 'OPC.UA.DA.StructuredType' := '1'}
	sts					: ST_DosingProcessSimStatus;
END_VAR
VAR
	elapsed				: LREAL; //seconds since start, for the main flow swing
	
	//Timers
	deltaTime			: FB_DeltaTime; //scan time
END_VAR
VAR CONSTANT
	TWO_PI				: LREAL := 6.283185307179586;
END_VAR

IF NOT cfg.enable THEN
	RETURN;
END_IF

Simulate();

METHOD PROTECTED Simulate
VAR
	period	: LREAL; //swing period in s
	lag		: LREAL; //process lag in s
END_VAR
deltaTime();
elapsed := elapsed + deltaTime.seconds;
period := TIME_TO_LREAL(cfg.swingPeriod) / 1000.0;
lag := TIME_TO_LREAL(cfg.processLag) / 1000.0;

//Main flow: slow swing around the base value
IF period > 0 THEN
	sts.mainFlow := cfg.mainFlowBase + cfg.mainFlowSwing * SIN(TWO_PI * elapsed / period);
ELSE
	sts.mainFlow := cfg.mainFlowBase;
END_IF

//Dosing flow: follows the valve position with a first-order lag
sts.dosingFlow := sts.dosingFlow + deltaTime.seconds / (lag + deltaTime.seconds)
				* (station.dosingValve.sts.position / 100.0 * cfg.maxDosingFlow - sts.dosingFlow);

station.flowMain.ctrl.sim := TRUE;
station.flowMain.ctrl.simValue := sts.mainFlow;
station.flowDosing.ctrl.sim := TRUE;
station.flowDosing.ctrl.simValue := sts.dosingFlow;
END_METHOD

END_FUNCTION_BLOCK
